// TIA Portal V17 program export: 0 tag tables, 0 data types, 1 data blocks, 1 code blocks (in call order from the OBs), 0 instance data blocks

DATA_BLOCK "AnimationTimer"   // DB1
{ S7_Optimized_Access := 'FALSE' }
   VAR
      T1 : TON_TIME;
      T2 : TON_TIME;
      T3 : TON_TIME;
      T4 : TON_TIME;
   END_VAR
BEGIN
END_DATA_BLOCK

ORGANIZATION_BLOCK "Main"   // OB1, LAD, ProgramCycle
TITLE = "Main Program Sweep (Cycle)"
{ S7_Optimized_Access := 'TRUE' }
// Codex 通过 V17 Openness 导入的原生 LAD 仿真示例。
// stored: SetENOAutomatically false
   VAR_INPUT
      Initial_Call : Bool;   // Initial call of this OB
      Remanence : Bool;   // =True, if remanent data are available
   END_VAR
BEGIN

REGION Network 1: 动画时基
   // 定时器每125毫秒产生一个扫描周期的脉冲。
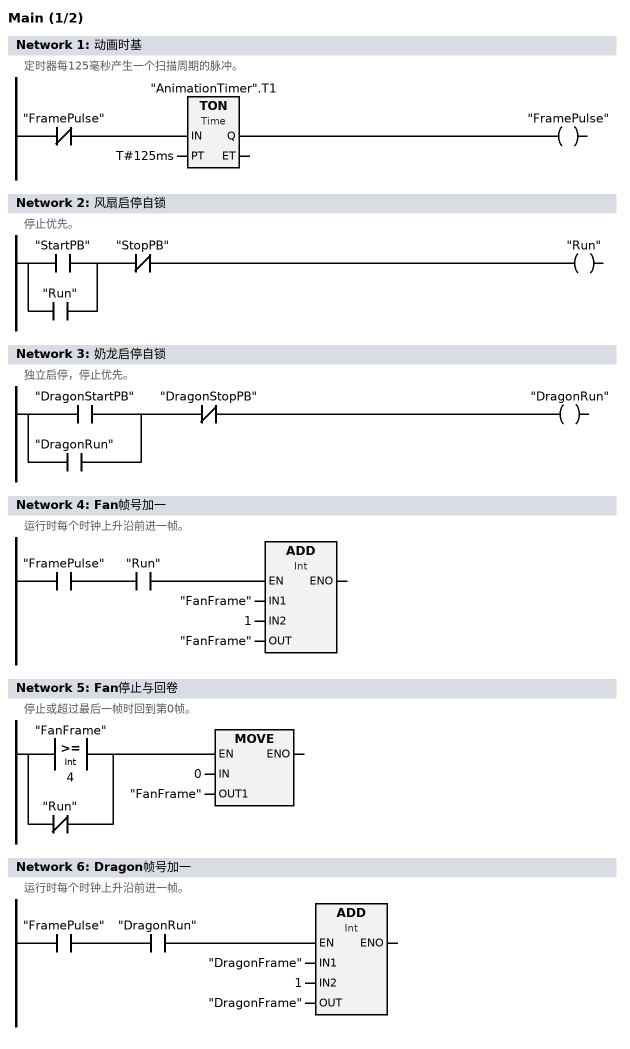
   RUNG wire#powerrail
      I_Contact( "FramePulse" )
      { S7_Templates := "time_type := Time" } "AnimationTimer".T1.TON(pt := T#125ms, et =>)
      Coil( "FramePulse" )
   END_RUNG
   // the same network as SCL:
   "AnimationTimer".T1.TON(IN := NOT "FramePulse", PT := T#125ms);
   "FramePulse" := "AnimationTimer".T1.Q;
END_REGION

REGION Network 2: 风扇启停自锁
   // 停止优先。
   RUNG wire#powerrail
      Contact( "StartPB" )
      wire#w1
      I_Contact( "StopPB" )
      Coil( "Run" )
   END_RUNG
   RUNG wire#powerrail
      Contact( "Run" )
   END_RUNG wire#w1
   // the same network as SCL:
   "Run" := ("StartPB" OR "Run") AND NOT "StopPB";
END_REGION

REGION Network 3: 奶龙启停自锁
   // 独立启停，停止优先。
   RUNG wire#powerrail
      Contact( "DragonStartPB" )
      wire#w1
      I_Contact( "DragonStopPB" )
      Coil( "DragonRun" )
   END_RUNG
   RUNG wire#powerrail
      Contact( "DragonRun" )
   END_RUNG wire#w1
   // the same network as SCL:
   "DragonRun" := ("DragonStartPB" OR "DragonRun") AND NOT "DragonStopPB";
END_REGION

REGION Network 4: Fan帧号加一
   // 运行时每个时钟上升沿前进一帧。
   RUNG wire#powerrail
      Contact( "FramePulse" )
      Contact( "Run" )
      { S7_Templates := "SrcType := Int" } Add(in1 := "FanFrame", in2 := 1, out := "FanFrame")
   END_RUNG
   // the same network as SCL:
   IF "FramePulse" AND "Run" THEN <??.?> := "FanFrame" + 1 + "FanFrame"; END_IF;
END_REGION

REGION Network 5: Fan停止与回卷
   // 停止或超过最后一帧时回到第0帧。
   RUNG wire#powerrail
      { S7_Templates := "SrcType := Int" } GE_Contact(in1 := "FanFrame", in2 := 4)
      wire#w1
      Move(in := 0, out1 := "FanFrame")
   END_RUNG
   RUNG wire#powerrail
      I_Contact( "Run" )
   END_RUNG wire#w1
   // the same network as SCL:
   IF ("FanFrame" >= 4) OR NOT "Run" THEN <??.?> := 0; END_IF;
END_REGION

REGION Network 6: Dragon帧号加一
   // 运行时每个时钟上升沿前进一帧。
   RUNG wire#powerrail
      Contact( "FramePulse" )
      Contact( "DragonRun" )
      { S7_Templates := "SrcType := Int" } Add(in1 := "DragonFrame", in2 := 1, out := "DragonFrame")
   END_RUNG
   // the same network as SCL:
   IF "FramePulse" AND "DragonRun" THEN <??.?> := "DragonFrame" + 1 + "DragonFrame"; END_IF;
END_REGION

REGION Network 7: Dragon停止与回卷
   // 停止或超过最后一帧时回到第0帧。
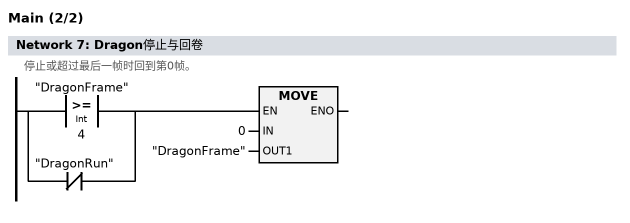
   RUNG wire#powerrail
      { S7_Templates := "SrcType := Int" } GE_Contact(in1 := "DragonFrame", in2 := 4)
      wire#w1
      Move(in := 0, out1 := "DragonFrame")
   END_RUNG
   RUNG wire#powerrail
      I_Contact( "DragonRun" )
   END_RUNG wire#w1
   // the same network as SCL:
   IF ("DragonFrame" >= 4) OR NOT "DragonRun" THEN <??.?> := 0; END_IF;
END_REGION
END_ORGANIZATION_BLOCK
